Fanuc KAREL source: kb00031.KL

PROGRAM KB00031
%STACKSIZE=65535
%PRIORITY=65535
%NOLOCKGROUP
VAR
P1 : REAL
P2 : STRING[80]
P3 : INTEGER
BEGIN
P1=1.0
P2='A'
P3=1
CNC_DYN_DISR(P1,P2,P3)
END KB00031
